(* Logix 5000 project; controller CIP_14485201 vendor 1 type 14 code 216 rev 38.11; software revision 38.01; part 8 of 12 *)
(* tags used below, declared in another part *)
   MOA_Drain_Flow_Mod_Value_Ind : INT;   // PV DRAIN FLOW MODULATION VALUE STATUS
   MOA_OFF : DINT[20];   // PANELVIEW MOA OFF
   MOA_ON : DINT[20];   // PANELVIEW MOA ON
   Panelview : INT[40];   // PANELVIEW CONTROL
   PV_Output_Status : INT[20];   // PV OUTPUT STATUS:
   PV_Output_Status_IND : INT[20,16];   // PV OUTPUT STATUS IND:
   PV_Status_Bit : BOOL;   // SYSTEM BIT
   SP_Drain_Flow : REAL;   // CURRENT DRAIN FLOW MODULATION SETPOINT
   Time_Date : DINT[20];   // SYSTEM TIME/DATE EDIT/STORAGE
(* MainProgram, continued *)

ROUTINE _07_SCALING   (* function block diagram *)
   SHEET 1   // Analog Input Scaling
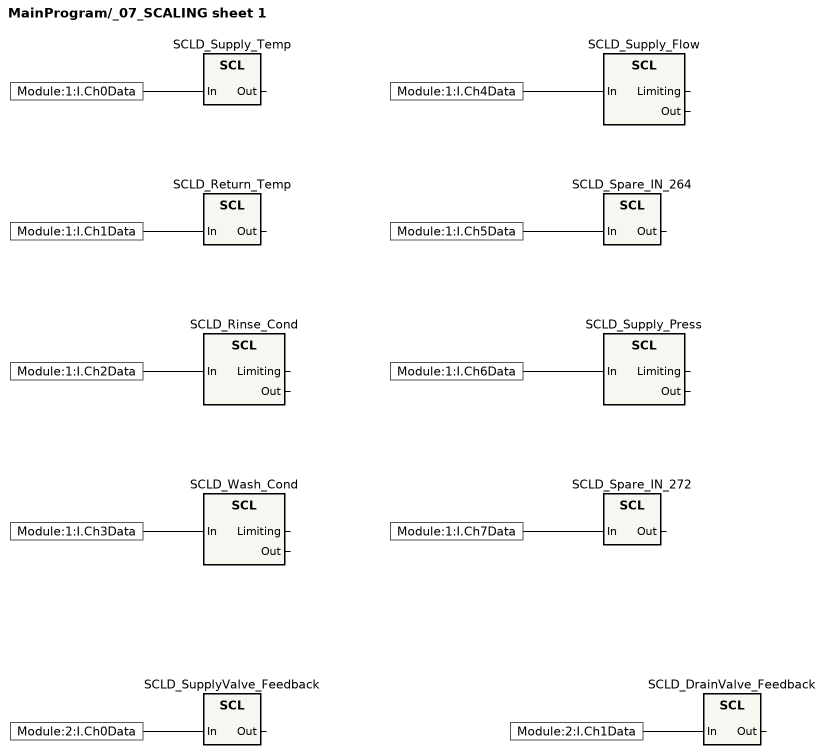
   SCLD_Supply_Temp : SCL(In := Module:1:I.Ch0Data);   // unwired pins: Out
   SCLD_Return_Temp : SCL(In := Module:1:I.Ch1Data);   // unwired pins: Out
   SCLD_Rinse_Cond : SCL(In := Module:1:I.Ch2Data);   // unwired pins: Limiting Out
   SCLD_Wash_Cond : SCL(In := Module:1:I.Ch3Data);   // unwired pins: Limiting Out
   SCLD_SupplyValve_Feedback : SCL(In := Module:2:I.Ch0Data);   // unwired pins: Out
   SCLD_Supply_Flow : SCL(In := Module:1:I.Ch4Data);   // unwired pins: Limiting Out
   SCLD_Spare_IN_264 : SCL(In := Module:1:I.Ch5Data);   // unwired pins: Out
   SCLD_Supply_Press : SCL(In := Module:1:I.Ch6Data);   // unwired pins: Limiting Out
   SCLD_Spare_IN_272 : SCL(In := Module:1:I.Ch7Data);   // unwired pins: Out
   SCLD_DrainValve_Feedback : SCL(In := Module:2:I.Ch1Data);   // unwired pins: Out
   SHEET 2   // Analog Output Scaling
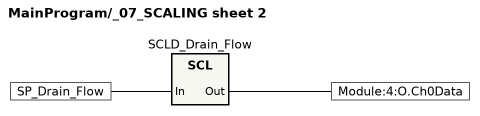
   SCLD_Drain_Flow : SCL(In := SP_Drain_Flow);
   Module:4:O.Ch0Data := SCLD_Drain_Flow.Out;
END_ROUTINE

ROUTINE _100_PV_STATUS   (* ladder *)
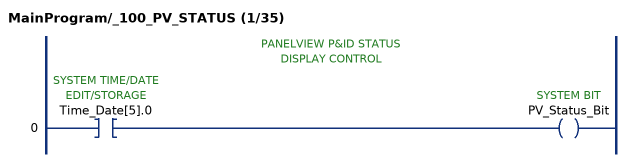
   // PANELVIEW P&ID STATUS
   // DISPLAY CONTROL
   0: XIC(Time_Date[5].0)OTE(PV_Status_Bit);
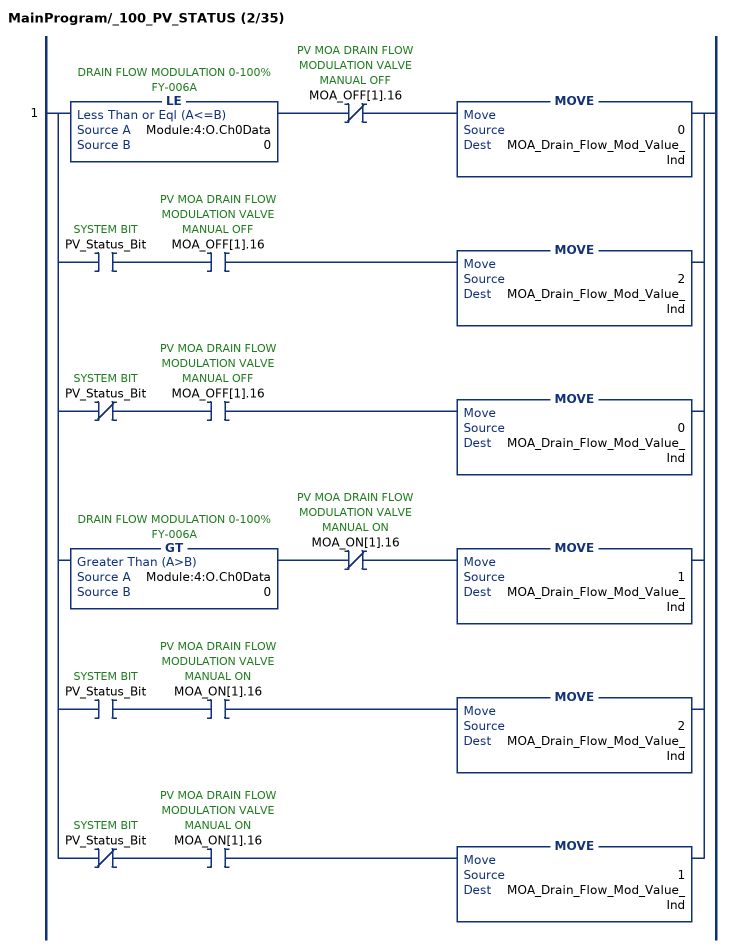
   1: [[LE(Module:4:O.Ch0Data,0) XIO(MOA_OFF[1].16) MOVE(0,MOA_Drain_Flow_Mod_Value_Ind) ,XIC(PV_Status_Bit) XIC(MOA_OFF[1].16) MOVE(2,MOA_Drain_Flow_Mod_Value_Ind) ,XIO(PV_Status_Bit) XIC(MOA_OFF[1].16) MOVE(0,MOA_Drain_Flow_Mod_Value_Ind) ] ,[GT(Module:4:O.Ch0Data,0) XIO(MOA_ON[1].16) MOVE(1,MOA_Drain_Flow_Mod_Value_Ind) ,XIC(PV_Status_Bit) XIC(MOA_ON[1].16) MOVE(2,MOA_Drain_Flow_Mod_Value_Ind) ,XIO(PV_Status_Bit) XIC(MOA_ON[1].16) MOVE(1,MOA_Drain_Flow_Mod_Value_Ind) ] ];
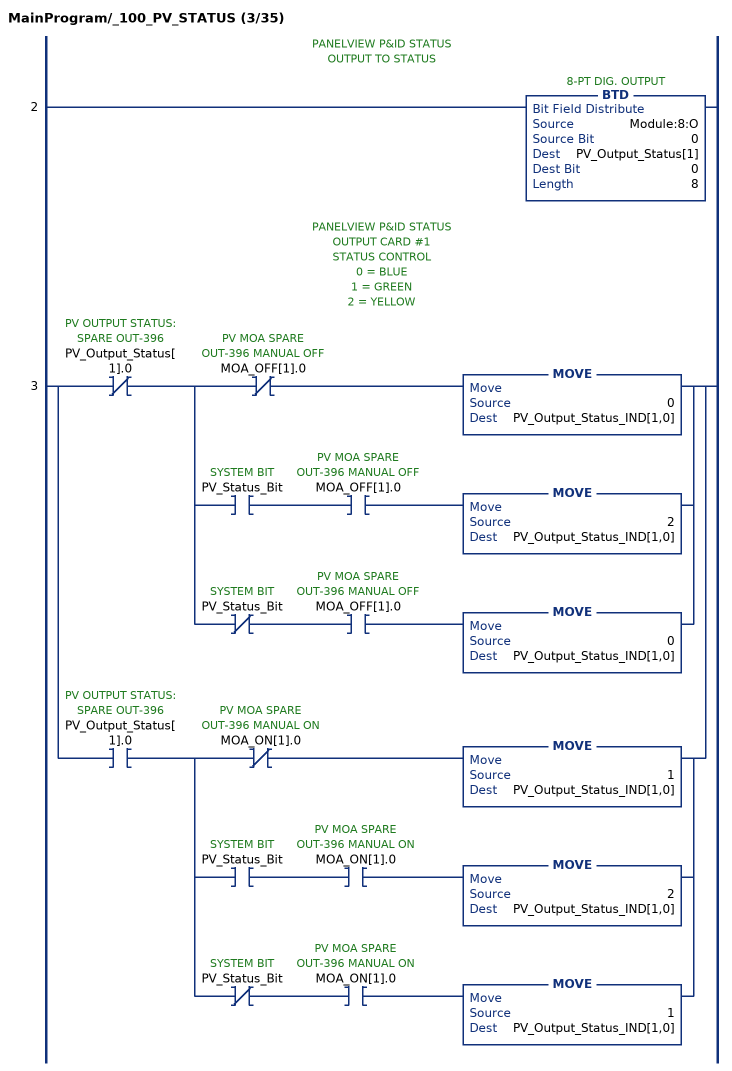
   // PANELVIEW P&ID STATUS
   // OUTPUT TO STATUS
   2: BTD(Module:8:O,0,PV_Output_Status[1],0,8);
   // PANELVIEW P&ID STATUS
   // OUTPUT CARD #1
   // STATUS CONTROL
   // 0 = BLUE
   // 1 = GREEN
   // 2 = YELLOW
   3: [XIO(PV_Output_Status[1].0) [XIO(MOA_OFF[1].0) MOVE(0,PV_Output_Status_IND[1,0]) ,XIC(PV_Status_Bit) XIC(MOA_OFF[1].0) MOVE(2,PV_Output_Status_IND[1,0]) ,XIO(PV_Status_Bit) XIC(MOA_OFF[1].0) MOVE(0,PV_Output_Status_IND[1,0]) ] ,XIC(PV_Output_Status[1].0) [XIO(MOA_ON[1].0) MOVE(1,PV_Output_Status_IND[1,0]) ,XIC(PV_Status_Bit) XIC(MOA_ON[1].0) MOVE(2,PV_Output_Status_IND[1,0]) ,XIO(PV_Status_Bit) XIC(MOA_ON[1].0) MOVE(1,PV_Output_Status_IND[1,0]) ] ];
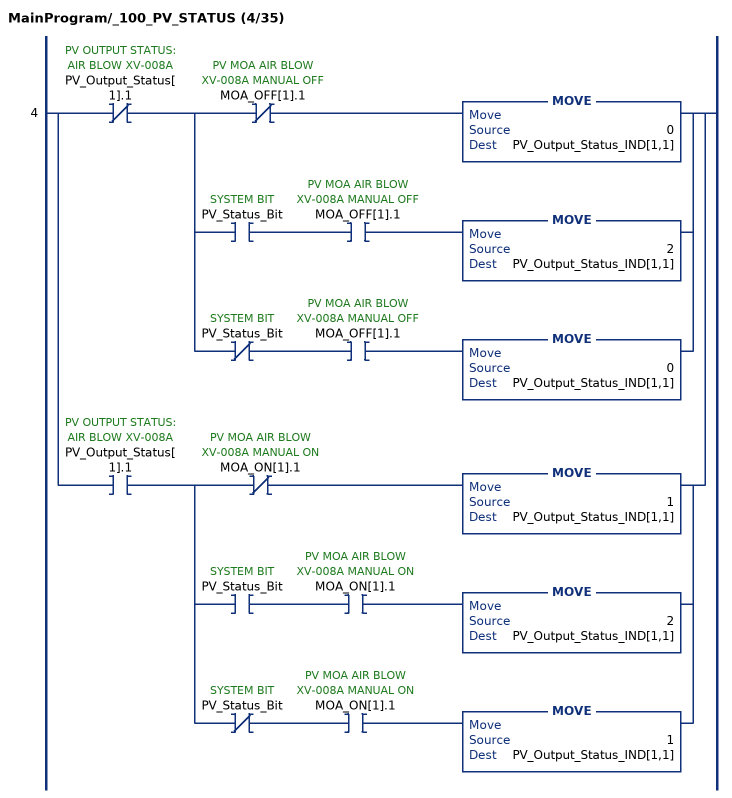
   4: [XIO(PV_Output_Status[1].1) [XIO(MOA_OFF[1].1) MOVE(0,PV_Output_Status_IND[1,1]) ,XIC(PV_Status_Bit) XIC(MOA_OFF[1].1) MOVE(2,PV_Output_Status_IND[1,1]) ,XIO(PV_Status_Bit) XIC(MOA_OFF[1].1) MOVE(0,PV_Output_Status_IND[1,1]) ] ,XIC(PV_Output_Status[1].1) [XIO(MOA_ON[1].1) MOVE(1,PV_Output_Status_IND[1,1]) ,XIC(PV_Status_Bit) XIC(MOA_ON[1].1) MOVE(2,PV_Output_Status_IND[1,1]) ,XIO(PV_Status_Bit) XIC(MOA_ON[1].1) MOVE(1,PV_Output_Status_IND[1,1]) ] ];
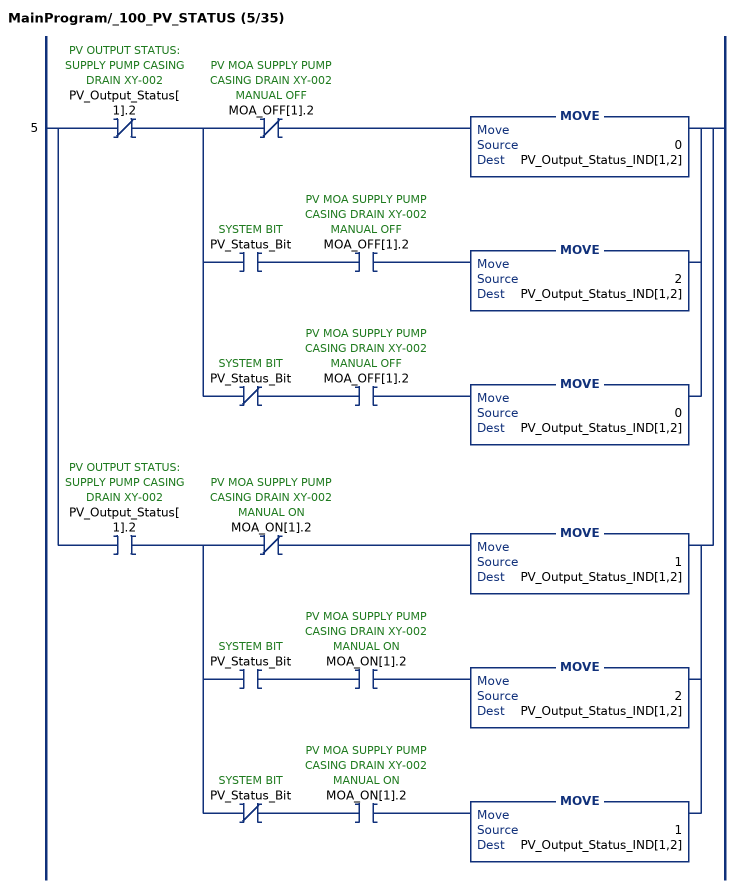
   5: [XIO(PV_Output_Status[1].2) [XIO(MOA_OFF[1].2) MOVE(0,PV_Output_Status_IND[1,2]) ,XIC(PV_Status_Bit) XIC(MOA_OFF[1].2) MOVE(2,PV_Output_Status_IND[1,2]) ,XIO(PV_Status_Bit) XIC(MOA_OFF[1].2) MOVE(0,PV_Output_Status_IND[1,2]) ] ,XIC(PV_Output_Status[1].2) [XIO(MOA_ON[1].2) MOVE(1,PV_Output_Status_IND[1,2]) ,XIC(PV_Status_Bit) XIC(MOA_ON[1].2) MOVE(2,PV_Output_Status_IND[1,2]) ,XIO(PV_Status_Bit) XIC(MOA_ON[1].2) MOVE(1,PV_Output_Status_IND[1,2]) ] ];
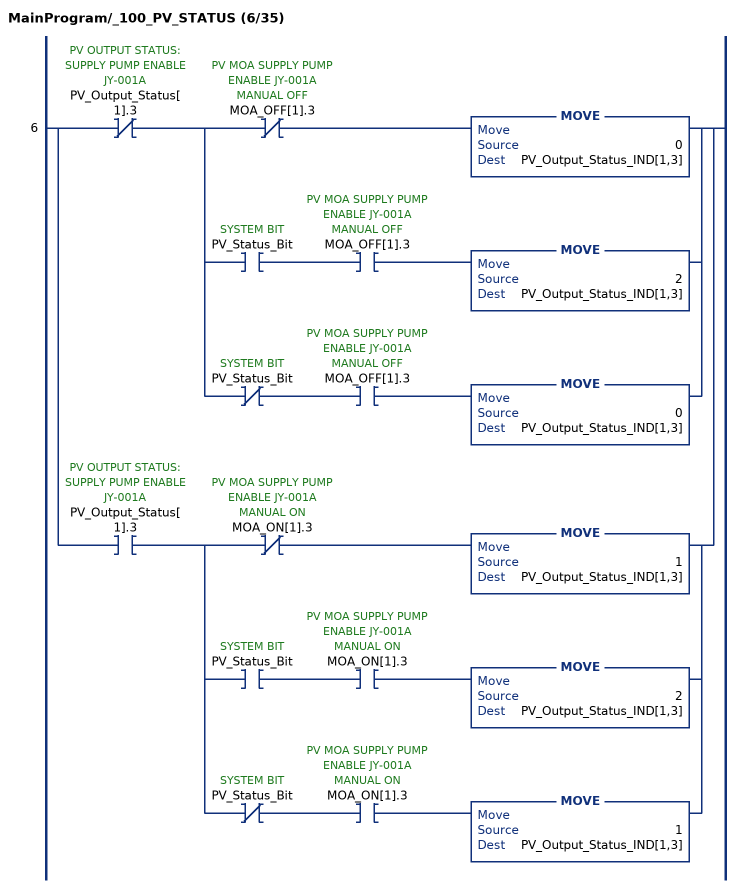
   6: [XIO(PV_Output_Status[1].3) [XIO(MOA_OFF[1].3) MOVE(0,PV_Output_Status_IND[1,3]) ,XIC(PV_Status_Bit) XIC(MOA_OFF[1].3) MOVE(2,PV_Output_Status_IND[1,3]) ,XIO(PV_Status_Bit) XIC(MOA_OFF[1].3) MOVE(0,PV_Output_Status_IND[1,3]) ] ,XIC(PV_Output_Status[1].3) [XIO(MOA_ON[1].3) MOVE(1,PV_Output_Status_IND[1,3]) ,XIC(PV_Status_Bit) XIC(MOA_ON[1].3) MOVE(2,PV_Output_Status_IND[1,3]) ,XIO(PV_Status_Bit) XIC(MOA_ON[1].3) MOVE(1,PV_Output_Status_IND[1,3]) ] ];
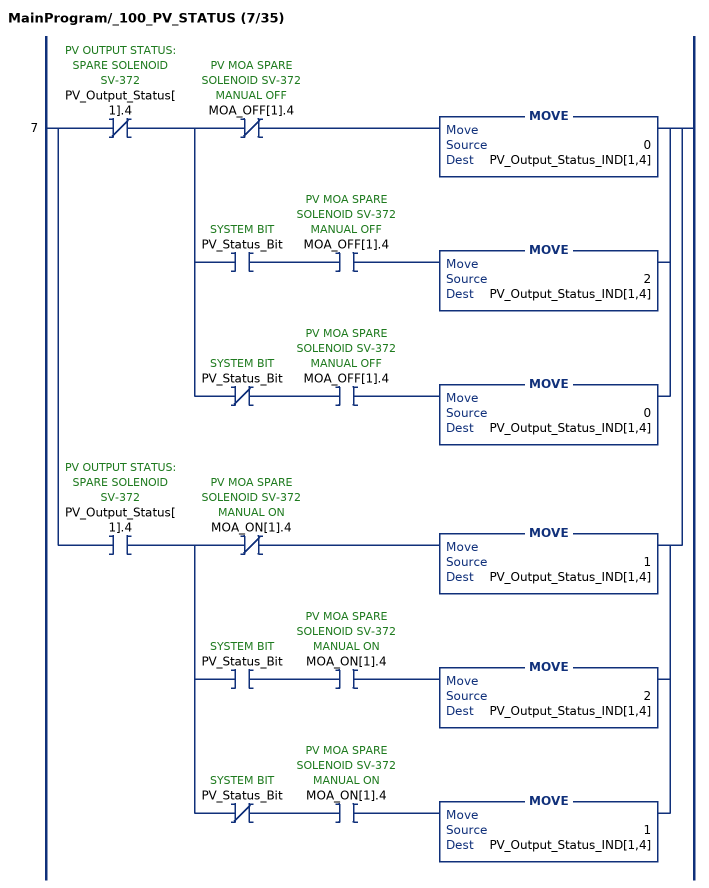
   7: [XIO(PV_Output_Status[1].4) [XIO(MOA_OFF[1].4) MOVE(0,PV_Output_Status_IND[1,4]) ,XIC(PV_Status_Bit) XIC(MOA_OFF[1].4) MOVE(2,PV_Output_Status_IND[1,4]) ,XIO(PV_Status_Bit) XIC(MOA_OFF[1].4) MOVE(0,PV_Output_Status_IND[1,4]) ] ,XIC(PV_Output_Status[1].4) [XIO(MOA_ON[1].4) MOVE(1,PV_Output_Status_IND[1,4]) ,XIC(PV_Status_Bit) XIC(MOA_ON[1].4) MOVE(2,PV_Output_Status_IND[1,4]) ,XIO(PV_Status_Bit) XIC(MOA_ON[1].4) MOVE(1,PV_Output_Status_IND[1,4]) ] ];
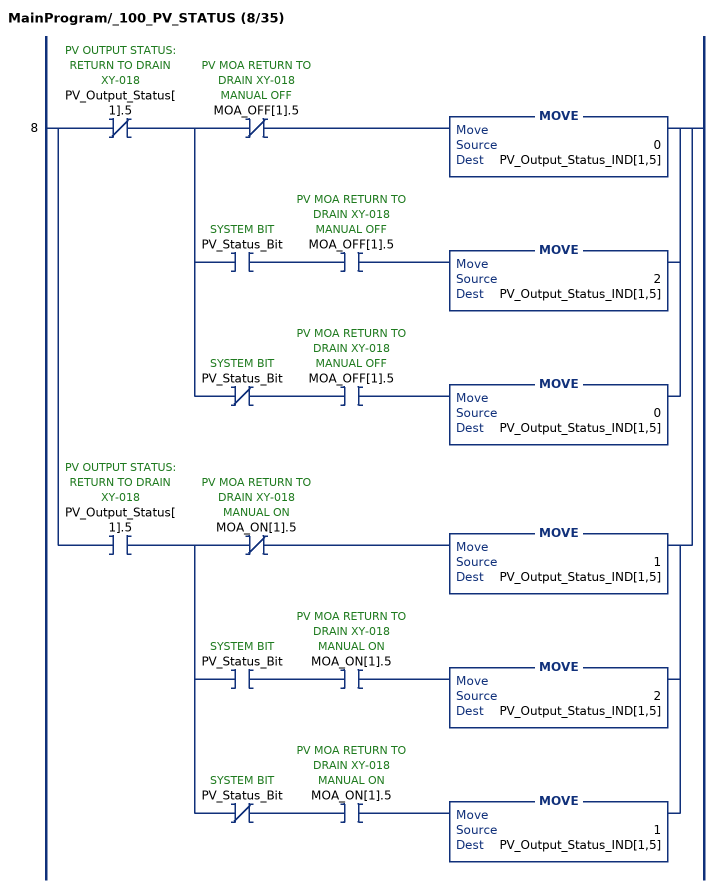
   8: [XIO(PV_Output_Status[1].5) [XIO(MOA_OFF[1].5) MOVE(0,PV_Output_Status_IND[1,5]) ,XIC(PV_Status_Bit) XIC(MOA_OFF[1].5) MOVE(2,PV_Output_Status_IND[1,5]) ,XIO(PV_Status_Bit) XIC(MOA_OFF[1].5) MOVE(0,PV_Output_Status_IND[1,5]) ] ,XIC(PV_Output_Status[1].5) [XIO(MOA_ON[1].5) MOVE(1,PV_Output_Status_IND[1,5]) ,XIC(PV_Status_Bit) XIC(MOA_ON[1].5) MOVE(2,PV_Output_Status_IND[1,5]) ,XIO(PV_Status_Bit) XIC(MOA_ON[1].5) MOVE(1,PV_Output_Status_IND[1,5]) ] ];
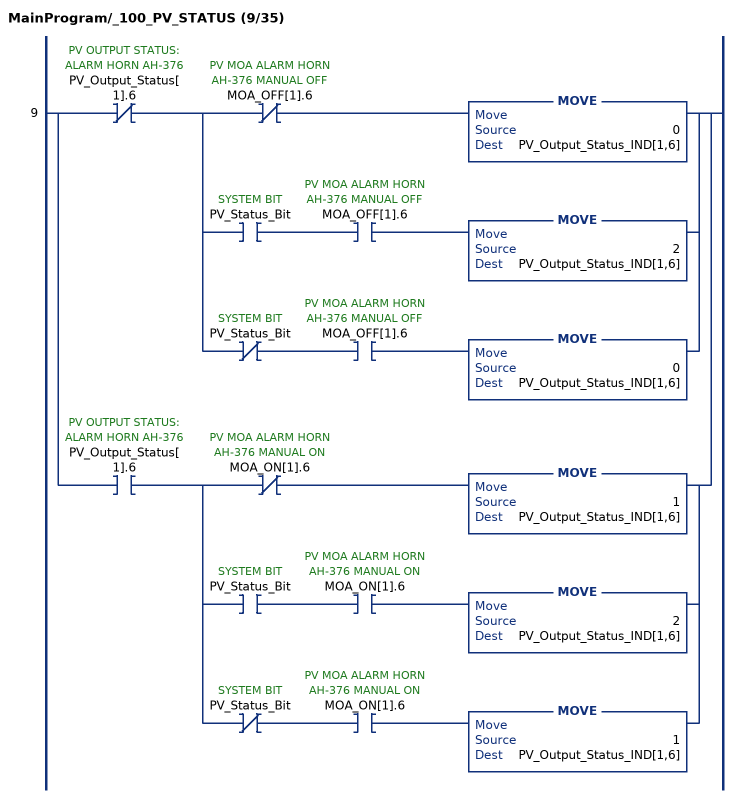
   9: [XIO(PV_Output_Status[1].6) [XIO(MOA_OFF[1].6) MOVE(0,PV_Output_Status_IND[1,6]) ,XIC(PV_Status_Bit) XIC(MOA_OFF[1].6) MOVE(2,PV_Output_Status_IND[1,6]) ,XIO(PV_Status_Bit) XIC(MOA_OFF[1].6) MOVE(0,PV_Output_Status_IND[1,6]) ] ,XIC(PV_Output_Status[1].6) [XIO(MOA_ON[1].6) MOVE(1,PV_Output_Status_IND[1,6]) ,XIC(PV_Status_Bit) XIC(MOA_ON[1].6) MOVE(2,PV_Output_Status_IND[1,6]) ,XIO(PV_Status_Bit) XIC(MOA_ON[1].6) MOVE(1,PV_Output_Status_IND[1,6]) ] ];
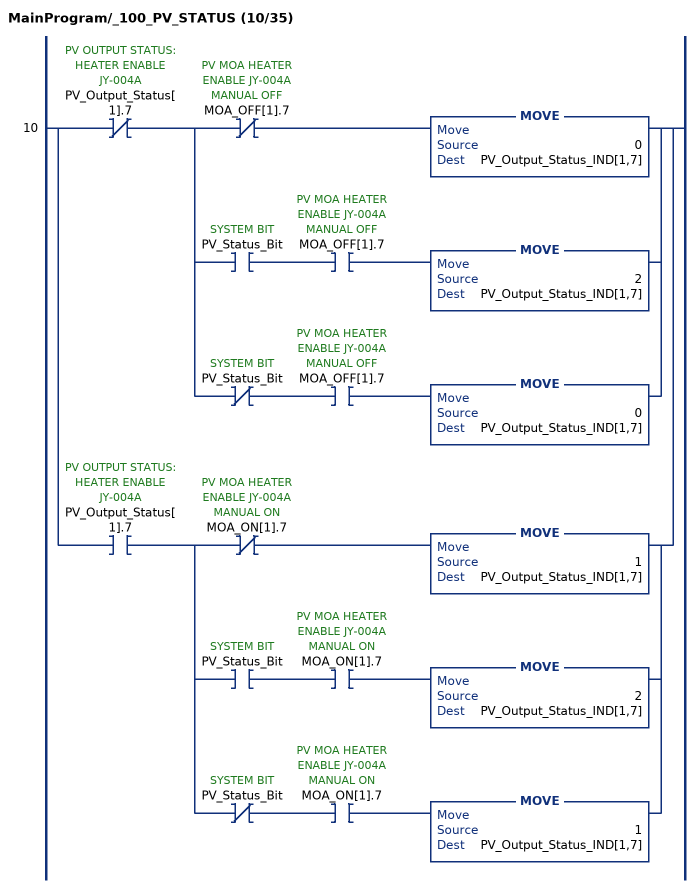
   10: [XIO(PV_Output_Status[1].7) [XIO(MOA_OFF[1].7) MOVE(0,PV_Output_Status_IND[1,7]) ,XIC(PV_Status_Bit) XIC(MOA_OFF[1].7) MOVE(2,PV_Output_Status_IND[1,7]) ,XIO(PV_Status_Bit) XIC(MOA_OFF[1].7) MOVE(0,PV_Output_Status_IND[1,7]) ] ,XIC(PV_Output_Status[1].7) [XIO(MOA_ON[1].7) MOVE(1,PV_Output_Status_IND[1,7]) ,XIC(PV_Status_Bit) XIC(MOA_ON[1].7) MOVE(2,PV_Output_Status_IND[1,7]) ,XIO(PV_Status_Bit) XIC(MOA_ON[1].7) MOVE(1,PV_Output_Status_IND[1,7]) ] ];
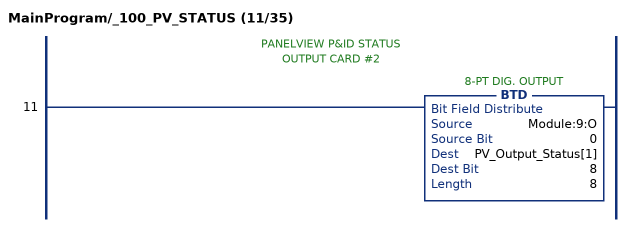
   // PANELVIEW P&ID STATUS
   // OUTPUT CARD #2
   11: BTD(Module:9:O,0,PV_Output_Status[1],8,8);
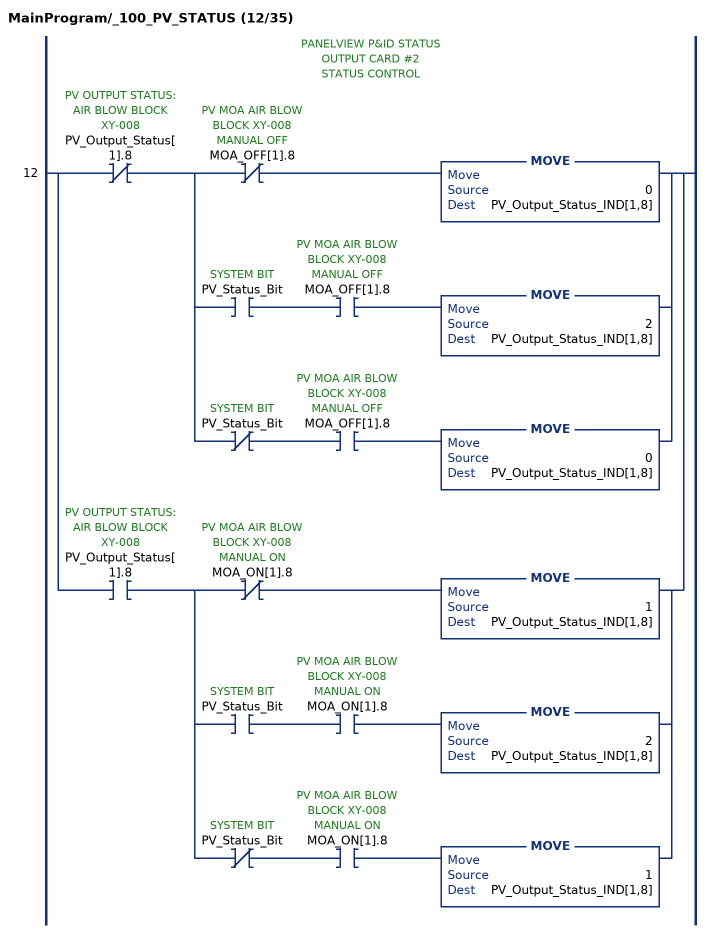
   // PANELVIEW P&ID STATUS
   // OUTPUT CARD #2
   // STATUS CONTROL
   12: [XIO(PV_Output_Status[1].8) [XIO(MOA_OFF[1].8) MOVE(0,PV_Output_Status_IND[1,8]) ,XIC(PV_Status_Bit) XIC(MOA_OFF[1].8) MOVE(2,PV_Output_Status_IND[1,8]) ,XIO(PV_Status_Bit) XIC(MOA_OFF[1].8) MOVE(0,PV_Output_Status_IND[1,8]) ] ,XIC(PV_Output_Status[1].8) [XIO(MOA_ON[1].8) MOVE(1,PV_Output_Status_IND[1,8]) ,XIC(PV_Status_Bit) XIC(MOA_ON[1].8) MOVE(2,PV_Output_Status_IND[1,8]) ,XIO(PV_Status_Bit) XIC(MOA_ON[1].8) MOVE(1,PV_Output_Status_IND[1,8]) ] ];
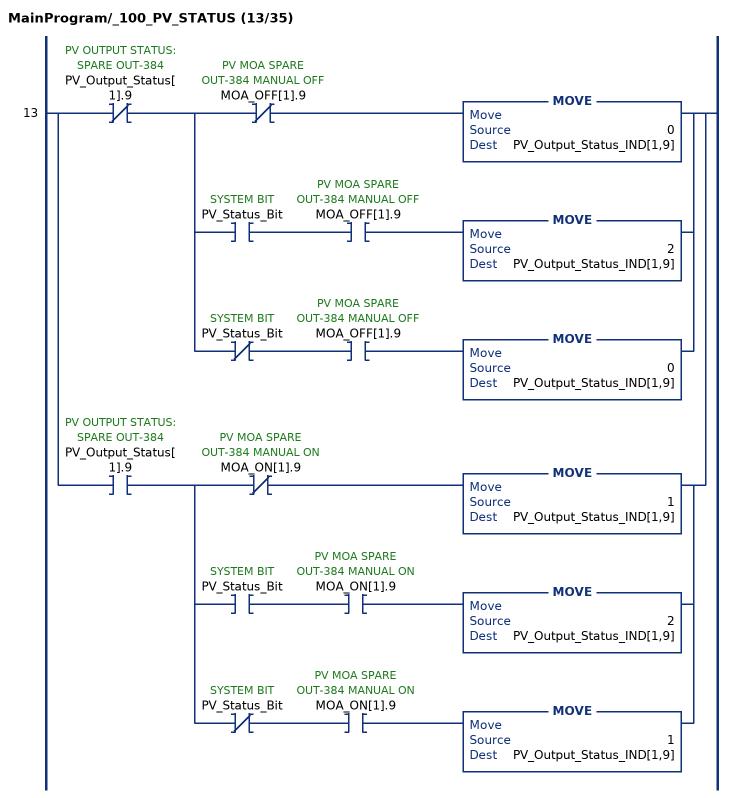
   13: [XIO(PV_Output_Status[1].9) [XIO(MOA_OFF[1].9) MOVE(0,PV_Output_Status_IND[1,9]) ,XIC(PV_Status_Bit) XIC(MOA_OFF[1].9) MOVE(2,PV_Output_Status_IND[1,9]) ,XIO(PV_Status_Bit) XIC(MOA_OFF[1].9) MOVE(0,PV_Output_Status_IND[1,9]) ] ,XIC(PV_Output_Status[1].9) [XIO(MOA_ON[1].9) MOVE(1,PV_Output_Status_IND[1,9]) ,XIC(PV_Status_Bit) XIC(MOA_ON[1].9) MOVE(2,PV_Output_Status_IND[1,9]) ,XIO(PV_Status_Bit) XIC(MOA_ON[1].9) MOVE(1,PV_Output_Status_IND[1,9]) ] ];
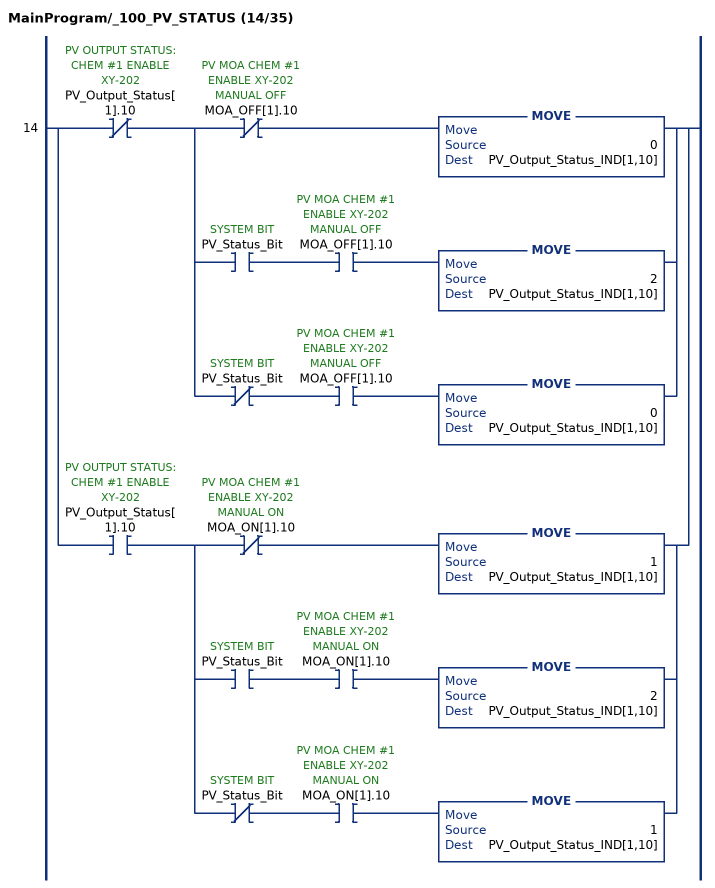
   14: [XIO(PV_Output_Status[1].10) [XIO(MOA_OFF[1].10) MOVE(0,PV_Output_Status_IND[1,10]) ,XIC(PV_Status_Bit) XIC(MOA_OFF[1].10) MOVE(2,PV_Output_Status_IND[1,10]) ,XIO(PV_Status_Bit) XIC(MOA_OFF[1].10) MOVE(0,PV_Output_Status_IND[1,10]) ] ,XIC(PV_Output_Status[1].10) [XIO(MOA_ON[1].10) MOVE(1,PV_Output_Status_IND[1,10]) ,XIC(PV_Status_Bit) XIC(MOA_ON[1].10) MOVE(2,PV_Output_Status_IND[1,10]) ,XIO(PV_Status_Bit) XIC(MOA_ON[1].10) MOVE(1,PV_Output_Status_IND[1,10]) ] ];
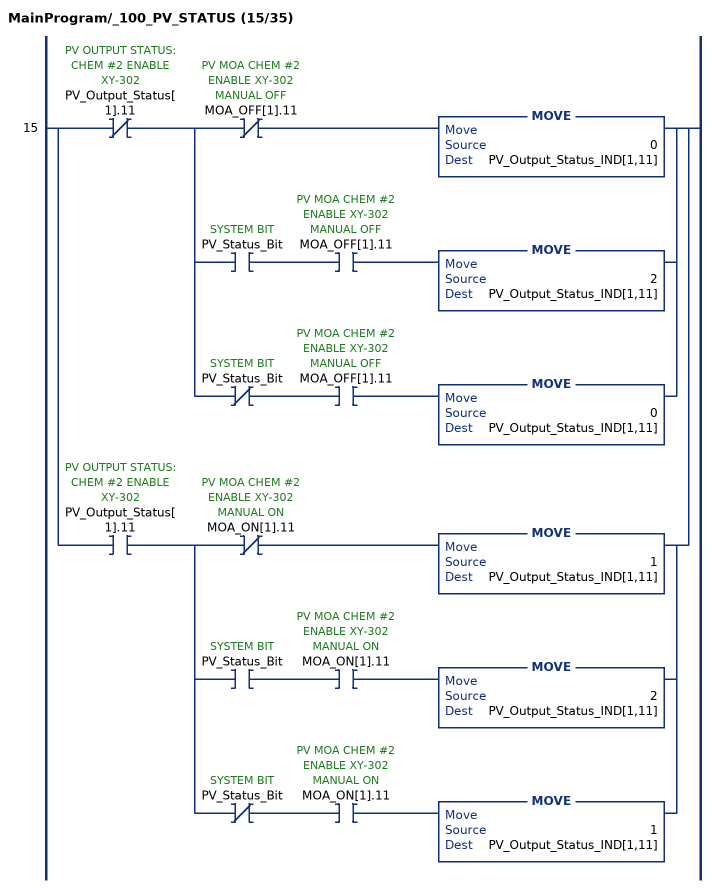
   15: [XIO(PV_Output_Status[1].11) [XIO(MOA_OFF[1].11) MOVE(0,PV_Output_Status_IND[1,11]) ,XIC(PV_Status_Bit) XIC(MOA_OFF[1].11) MOVE(2,PV_Output_Status_IND[1,11]) ,XIO(PV_Status_Bit) XIC(MOA_OFF[1].11) MOVE(0,PV_Output_Status_IND[1,11]) ] ,XIC(PV_Output_Status[1].11) [XIO(MOA_ON[1].11) MOVE(1,PV_Output_Status_IND[1,11]) ,XIC(PV_Status_Bit) XIC(MOA_ON[1].11) MOVE(2,PV_Output_Status_IND[1,11]) ,XIO(PV_Status_Bit) XIC(MOA_ON[1].11) MOVE(1,PV_Output_Status_IND[1,11]) ] ];
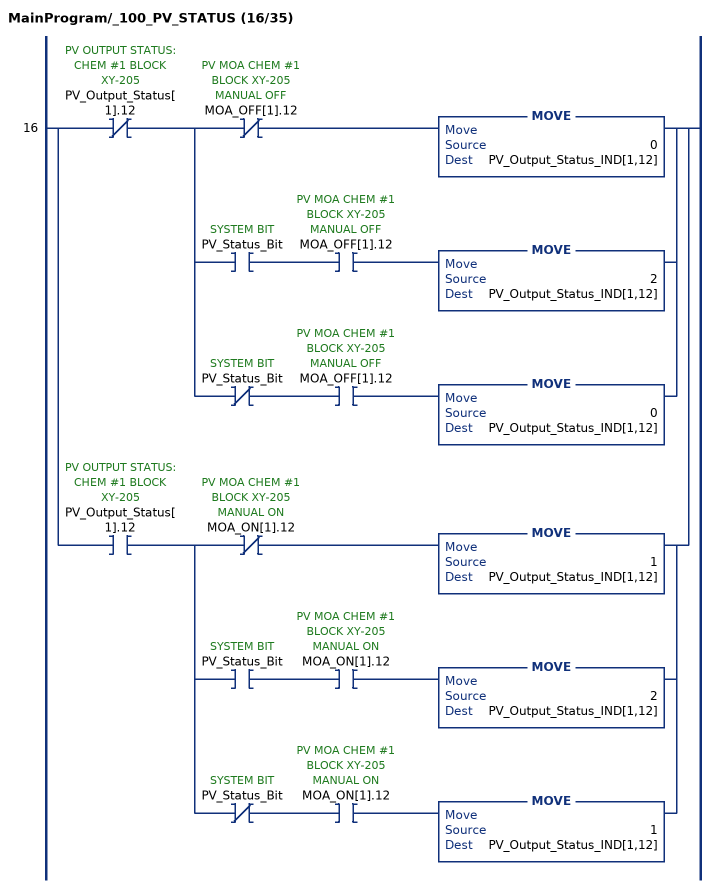
   16: [XIO(PV_Output_Status[1].12) [XIO(MOA_OFF[1].12) MOVE(0,PV_Output_Status_IND[1,12]) ,XIC(PV_Status_Bit) XIC(MOA_OFF[1].12) MOVE(2,PV_Output_Status_IND[1,12]) ,XIO(PV_Status_Bit) XIC(MOA_OFF[1].12) MOVE(0,PV_Output_Status_IND[1,12]) ] ,XIC(PV_Output_Status[1].12) [XIO(MOA_ON[1].12) MOVE(1,PV_Output_Status_IND[1,12]) ,XIC(PV_Status_Bit) XIC(MOA_ON[1].12) MOVE(2,PV_Output_Status_IND[1,12]) ,XIO(PV_Status_Bit) XIC(MOA_ON[1].12) MOVE(1,PV_Output_Status_IND[1,12]) ] ];
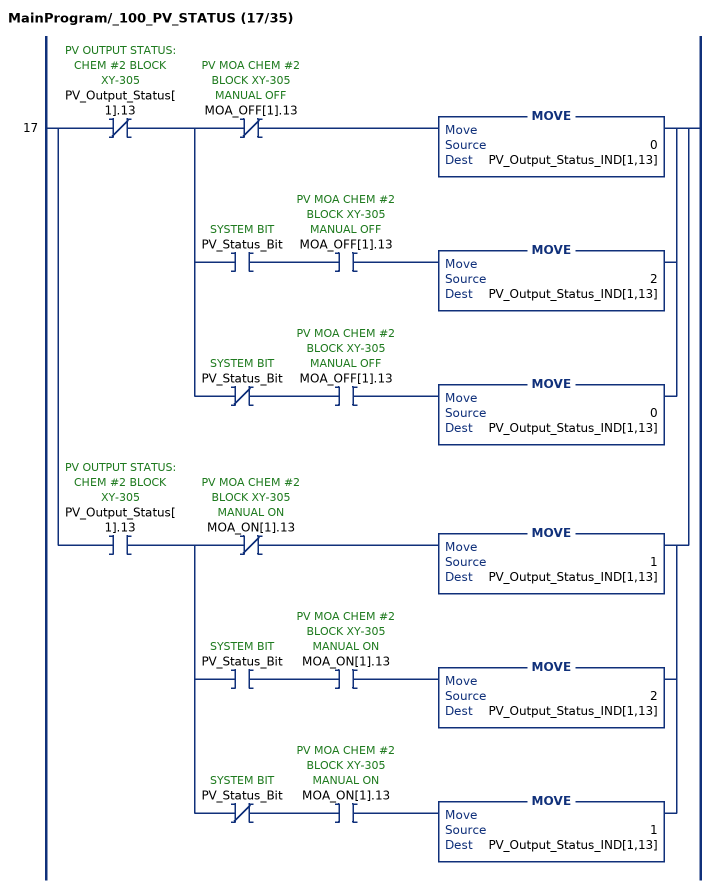
   17: [XIO(PV_Output_Status[1].13) [XIO(MOA_OFF[1].13) MOVE(0,PV_Output_Status_IND[1,13]) ,XIC(PV_Status_Bit) XIC(MOA_OFF[1].13) MOVE(2,PV_Output_Status_IND[1,13]) ,XIO(PV_Status_Bit) XIC(MOA_OFF[1].13) MOVE(0,PV_Output_Status_IND[1,13]) ] ,XIC(PV_Output_Status[1].13) [XIO(MOA_ON[1].13) MOVE(1,PV_Output_Status_IND[1,13]) ,XIC(PV_Status_Bit) XIC(MOA_ON[1].13) MOVE(2,PV_Output_Status_IND[1,13]) ,XIO(PV_Status_Bit) XIC(MOA_ON[1].13) MOVE(1,PV_Output_Status_IND[1,13]) ] ];
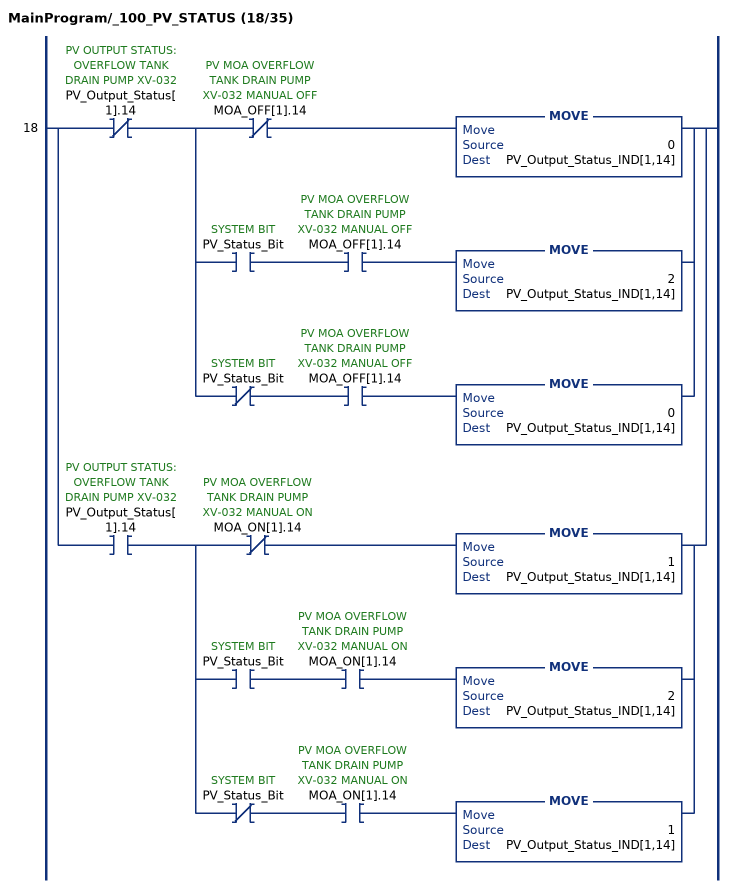
   18: [XIO(PV_Output_Status[1].14) [XIO(MOA_OFF[1].14) MOVE(0,PV_Output_Status_IND[1,14]) ,XIC(PV_Status_Bit) XIC(MOA_OFF[1].14) MOVE(2,PV_Output_Status_IND[1,14]) ,XIO(PV_Status_Bit) XIC(MOA_OFF[1].14) MOVE(0,PV_Output_Status_IND[1,14]) ] ,XIC(PV_Output_Status[1].14) [XIO(MOA_ON[1].14) MOVE(1,PV_Output_Status_IND[1,14]) ,XIC(PV_Status_Bit) XIC(MOA_ON[1].14) MOVE(2,PV_Output_Status_IND[1,14]) ,XIO(PV_Status_Bit) XIC(MOA_ON[1].14) MOVE(1,PV_Output_Status_IND[1,14]) ] ];
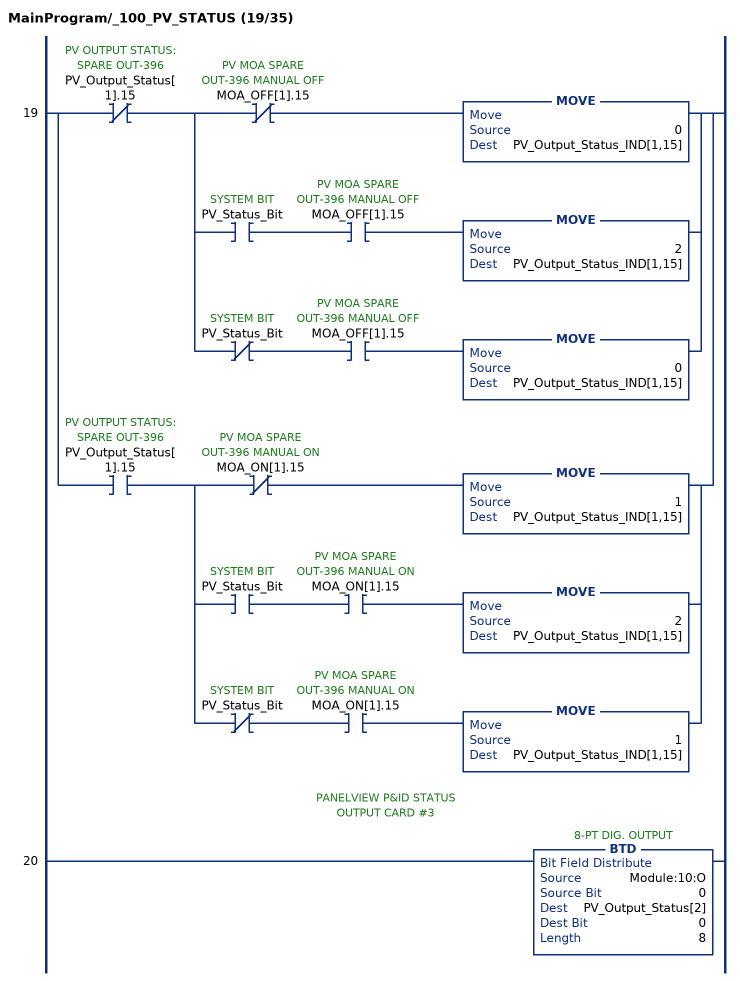
   19: [XIO(PV_Output_Status[1].15) [XIO(MOA_OFF[1].15) MOVE(0,PV_Output_Status_IND[1,15]) ,XIC(PV_Status_Bit) XIC(MOA_OFF[1].15) MOVE(2,PV_Output_Status_IND[1,15]) ,XIO(PV_Status_Bit) XIC(MOA_OFF[1].15) MOVE(0,PV_Output_Status_IND[1,15]) ] ,XIC(PV_Output_Status[1].15) [XIO(MOA_ON[1].15) MOVE(1,PV_Output_Status_IND[1,15]) ,XIC(PV_Status_Bit) XIC(MOA_ON[1].15) MOVE(2,PV_Output_Status_IND[1,15]) ,XIO(PV_Status_Bit) XIC(MOA_ON[1].15) MOVE(1,PV_Output_Status_IND[1,15]) ] ];
   // PANELVIEW P&ID STATUS
   // OUTPUT CARD #3
   20: BTD(Module:10:O,0,PV_Output_Status[2],0,8);
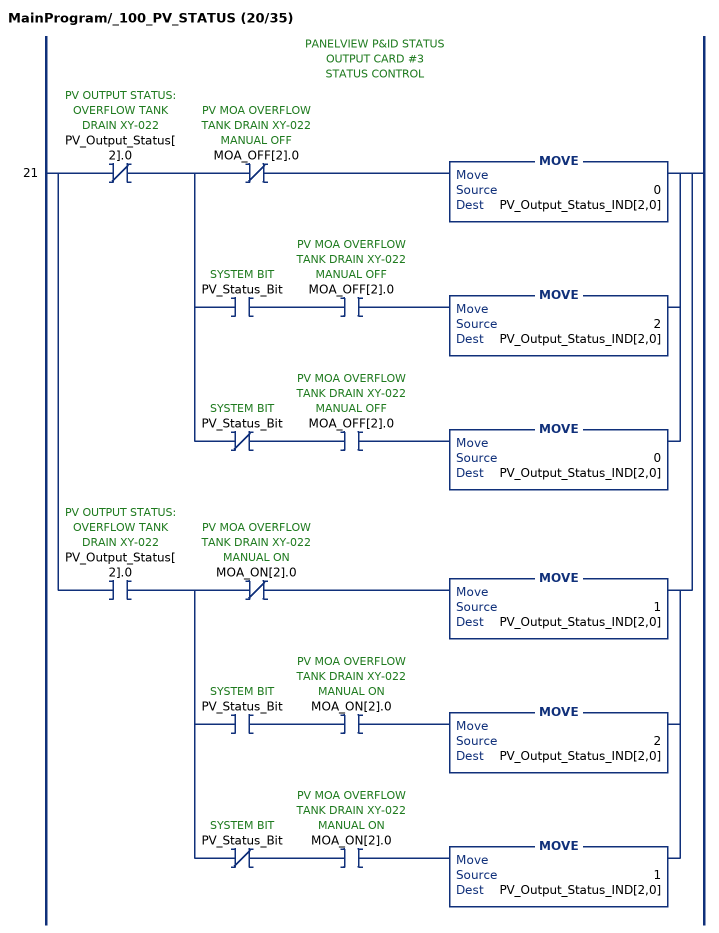
   // PANELVIEW P&ID STATUS
   // OUTPUT CARD #3
   // STATUS CONTROL
   21: [XIO(PV_Output_Status[2].0) [XIO(MOA_OFF[2].0) MOVE(0,PV_Output_Status_IND[2,0]) ,XIC(PV_Status_Bit) XIC(MOA_OFF[2].0) MOVE(2,PV_Output_Status_IND[2,0]) ,XIO(PV_Status_Bit) XIC(MOA_OFF[2].0) MOVE(0,PV_Output_Status_IND[2,0]) ] ,XIC(PV_Output_Status[2].0) [XIO(MOA_ON[2].0) MOVE(1,PV_Output_Status_IND[2,0]) ,XIC(PV_Status_Bit) XIC(MOA_ON[2].0) MOVE(2,PV_Output_Status_IND[2,0]) ,XIO(PV_Status_Bit) XIC(MOA_ON[2].0) MOVE(1,PV_Output_Status_IND[2,0]) ] ];
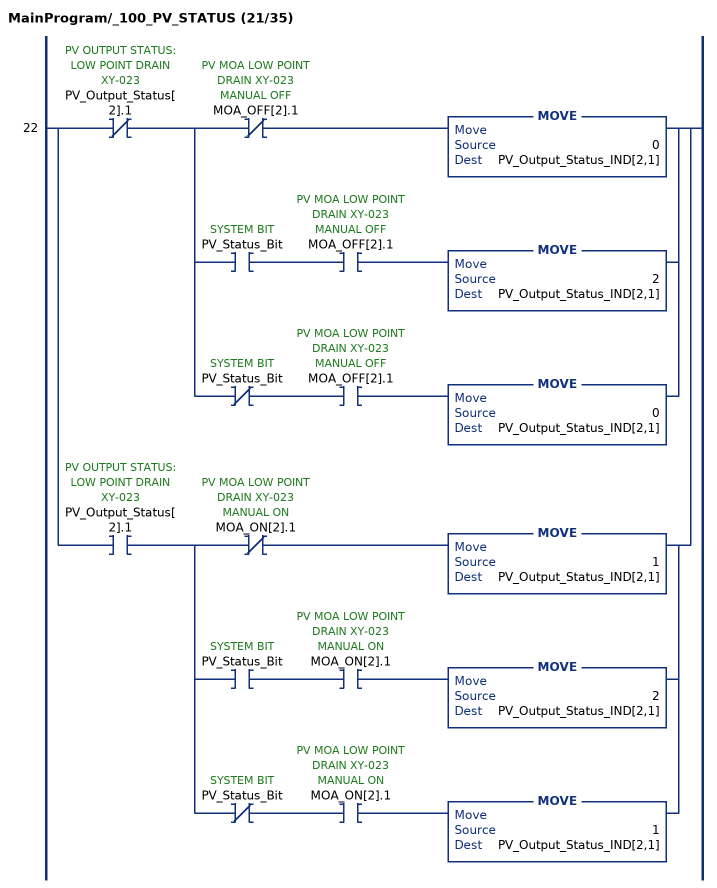
   22: [XIO(PV_Output_Status[2].1) [XIO(MOA_OFF[2].1) MOVE(0,PV_Output_Status_IND[2,1]) ,XIC(PV_Status_Bit) XIC(MOA_OFF[2].1) MOVE(2,PV_Output_Status_IND[2,1]) ,XIO(PV_Status_Bit) XIC(MOA_OFF[2].1) MOVE(0,PV_Output_Status_IND[2,1]) ] ,XIC(PV_Output_Status[2].1) [XIO(MOA_ON[2].1) MOVE(1,PV_Output_Status_IND[2,1]) ,XIC(PV_Status_Bit) XIC(MOA_ON[2].1) MOVE(2,PV_Output_Status_IND[2,1]) ,XIO(PV_Status_Bit) XIC(MOA_ON[2].1) MOVE(1,PV_Output_Status_IND[2,1]) ] ];
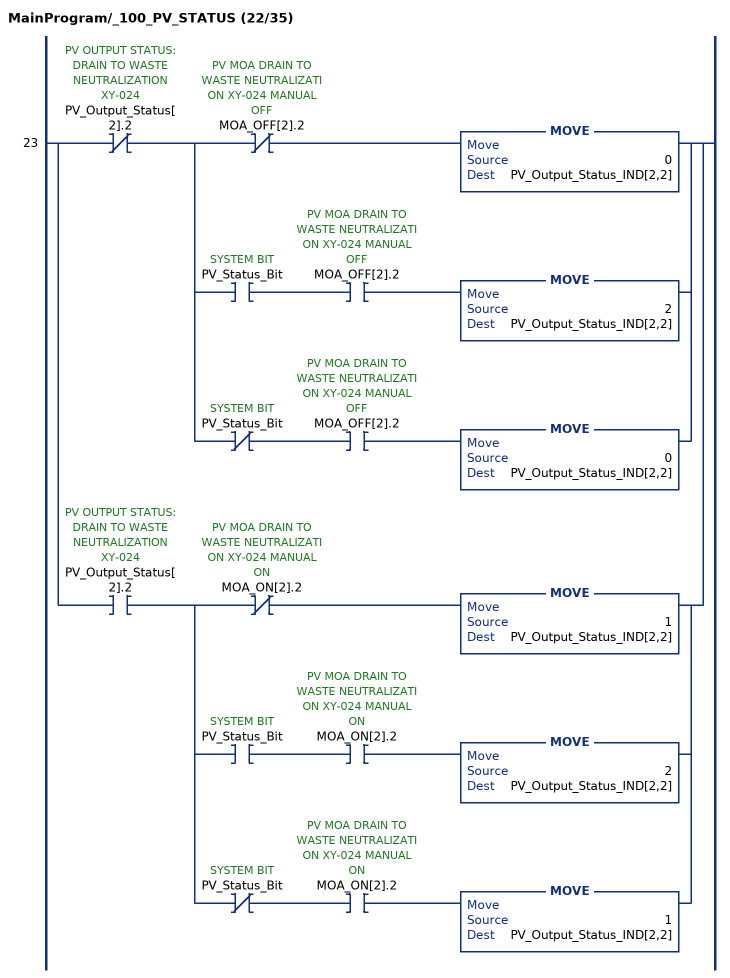
   23: [XIO(PV_Output_Status[2].2) [XIO(MOA_OFF[2].2) MOVE(0,PV_Output_Status_IND[2,2]) ,XIC(PV_Status_Bit) XIC(MOA_OFF[2].2) MOVE(2,PV_Output_Status_IND[2,2]) ,XIO(PV_Status_Bit) XIC(MOA_OFF[2].2) MOVE(0,PV_Output_Status_IND[2,2]) ] ,XIC(PV_Output_Status[2].2) [XIO(MOA_ON[2].2) MOVE(1,PV_Output_Status_IND[2,2]) ,XIC(PV_Status_Bit) XIC(MOA_ON[2].2) MOVE(2,PV_Output_Status_IND[2,2]) ,XIO(PV_Status_Bit) XIC(MOA_ON[2].2) MOVE(1,PV_Output_Status_IND[2,2]) ] ];
